// TIA Portal V21 export
// export: Created 2026-10-12T12:46:13.185712Z, ExportSetting WithDefaults, DisplayName Totally Integrated Automation Portal, DisplayVersion V21, DisplayName STEP 7 Professional, DisplayVersion V21, DisplayName STEP 7 Safety, DisplayVersion V21, DisplayName Tech WebApplication, DisplayVersion V21, DisplayName WinCC Basic/Comfort/Advanced, DisplayVersion V21, DisplayName WinCC Unified, DisplayVersion V21
Screen "AUTO"  800x480, Number=1, Template=MAIN
  ScreenLayer 
    TextField "Template_Text field_2" at 308,62 size 181x27  Text="AUTO OPERATION"
    SymbolicIOField "Symbolic I/O field_1" at 116,182 size 560x106  CountVisibleItems=3, Mode=Output, OnValue=1, TextList=AUTO STATUS, TextOff="0", TextOn="1"
      RangeAppearanceAnimation "RangeAppearanceAnimation"
        tag DB_AUTO_AUTO STATUS
        10..10: back #00ff00, fore #000000
        20..20: back #ff0000, fore #ffffff
      ProcessValue := DB_AUTO_AUTO STATUS
    TextField "Template_Text field_1" at 304,117 size 165x34  Text="AUTO STATUS"
